(* Logix 5000 project; controller Tank_Filling Emulate 5570 rev 33.11; software revision 33.03 *)
// Tank level control using Low Low, Low, High, and High High switches, with automatic filling, draining mode, and level alarms.

TASK MainTask (continuous, watchdog 500 ms) : MainProgram

MODULES
   Local : Emulate 5570 (ICP 3, rev 33.11)
END_MODULES

VAR_GLOBAL   (* controller tags *)
   Alarm_HH : BOOL;   // High high alarm
   Alarm_LL : BOOL;   // Low low alarm
   Alarm_Output : BOOL;   // Common alarm indicator
   Alarm_Reset : BOOL;   // Reset latched alarms
   Drain_Mode : BOOL;   // 0 = automatic filling; 1 = draining
   Drain_Output : BOOL;   // Drain pump or valve command
   Drain_Request : BOOL;   // Internal draining demand
   Fill_Request : BOOL;   // Internal filling demand
   HH_Alarm_Timer : TIMER := (PRE := 2000);
   Inlet_Output : BOOL;   // Inlet pump or valve command
   Level_H : BOOL;
   Level_HH : BOOL;
   Level_L : BOOL;
   Level_LL : BOOL;
   LL_Alarm_Timer : TIMER := (PRE := 2000);
   Reset_ONS : BOOL;
   Reset_Pulse : BOOL;
   Start_PB : BOOL;   // Start command
   Stop_Request : BOOL;   // Stop command: 1 = stop
   System_Run : BOOL;   // System enabled
END_VAR

PROGRAM MainProgram   (* main routine MainRoutine *)

ROUTINE MainRoutine   (* ladder *)
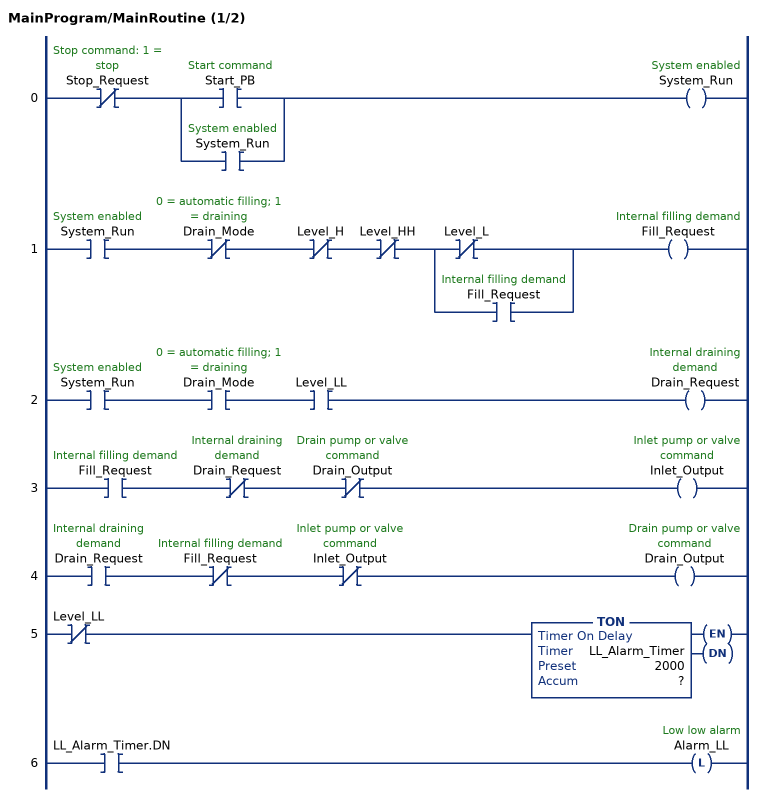
   0: XIO(Stop_Request)[XIC(Start_PB) ,XIC(System_Run) ]OTE(System_Run);
   1: XIC(System_Run)XIO(Drain_Mode)XIO(Level_H)XIO(Level_HH)[XIO(Level_L) ,XIC(Fill_Request) ]OTE(Fill_Request);
   2: XIC(System_Run)XIC(Drain_Mode)XIC(Level_LL)OTE(Drain_Request);
   3: XIC(Fill_Request)XIO(Drain_Request)XIO(Drain_Output)OTE(Inlet_Output);
   4: XIC(Drain_Request)XIO(Fill_Request)XIO(Inlet_Output)OTE(Drain_Output);
   5: XIO(Level_LL)TON(LL_Alarm_Timer,?,?);
   6: XIC(LL_Alarm_Timer.DN)OTL(Alarm_LL);
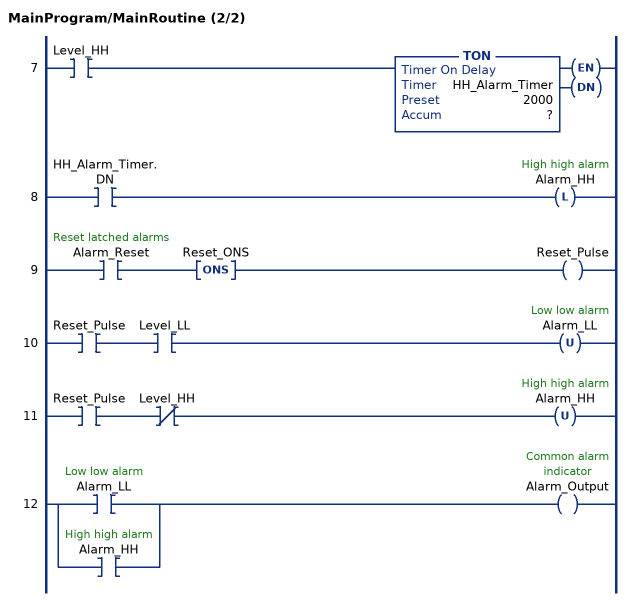
   7: XIC(Level_HH)TON(HH_Alarm_Timer,?,?);
   8: XIC(HH_Alarm_Timer.DN)OTL(Alarm_HH);
   9: XIC(Alarm_Reset)ONS(Reset_ONS)OTE(Reset_Pulse);
   10: XIC(Reset_Pulse)XIC(Level_LL)OTU(Alarm_LL);
   11: XIC(Reset_Pulse)XIO(Level_HH)OTU(Alarm_HH);
   12: [XIC(Alarm_LL) ,XIC(Alarm_HH) ]OTE(Alarm_Output);
END_ROUTINE
END_PROGRAM
